Fanuc KAREL source: KB00119.KL

PROGRAM KB00119
%NOLOCKGROUP
%ENVIRONMENT MULTI
VAR
  P1: INTEGER
  P2: INTEGER
BEGIN
  P1 = 1
  P2 = 1
  LOCK_GROUP(P1, P2)
END KB00119
